(*

**Autonumbered footnotes**

Autonumbered footnotes are possible, like using [#]_ and [#]_. 

--------

.. [#] This is the first one. 

.. [#] This is the second one. 
*)

FUNCTION_BLOCK FB_Libdoc_AutomaticallyNumberedFootnotes
VAR_INPUT
    nVarA : INT;
    nVarB : INT;
END_VAR
VAR_OUTPUT
    nSum : INT;
END_VAR
VAR
END_VAR

END_FUNCTION_BLOCK

(* stored: Version 1.1.0.1, ProductVersion 3.1.4022.17
   POU FB_Libdoc_AutomaticallyNumberedFootnotes: Id {8c689454-3d67-4efa-8828-810eb1f01367}, SpecialFunc None *)
